// SIMATIC STEP 7 (V5.x) project EXO6
// CPU: CPU 314
// station: Matériel
// station: SIMATIC 300(1)
// station: P_ADR_BUS
// program: Programme S7(1)

SYMBOL_TABLE
"BP"	I 0.0	BOOL
"MOTEUR"	Q 0.0	BOOL
"LAMPE"	Q 0.1	BOOL
END_SYMBOL_TABLE

ORGANIZATION_BLOCK OB 1
TITLE = "Main Program Sweep (Cycle)"
VERSION : 0.1
VAR_TEMP
  OB1_EV_CLASS : BYTE ;	//Bits 0-3 = 1 (Coming event), Bits 4-7 = 1 (Event class 1)
  OB1_SCAN_1 : BYTE ;	//1 (Cold restart scan 1 of OB 1), 3 (Scan 2-n of OB 1)
  OB1_PRIORITY : BYTE ;	//Priority of OB Execution
  OB1_OB_NUMBR : BYTE ;	//1 (Organization block 1, OB1)
  OB1_RESERVED_1 : BYTE ;	//Reserved for system
  OB1_RESERVED_2 : BYTE ;	//Reserved for system
  OB1_PREV_CYCLE : INT ;	//Cycle time of previous OB1 scan (milliseconds)
  OB1_MIN_CYCLE : INT ;	//Minimum cycle time of OB1 (milliseconds)
  OB1_MAX_CYCLE : INT ;	//Maximum cycle time of OB1 (milliseconds)
  OB1_DATE_TIME : DATE_AND_TIME ;	//Date and time OB1 started
END_VAR
BEGIN
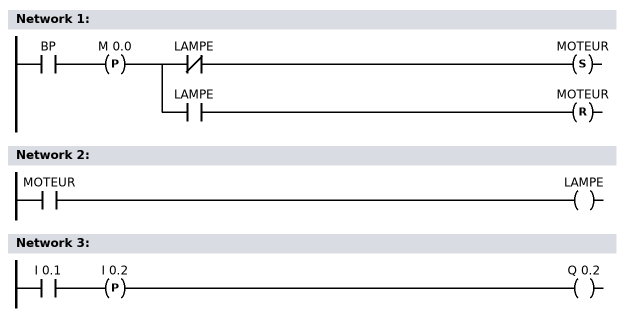
NETWORK
TITLE =
      A     "BP";
      BLD   100;
      FP    M 0.0;
      =     L 20.0;
      A     L 20.0;
      AN    "LAMPE";
      S     "MOTEUR";
      A     L 20.0;
      A     "LAMPE";
      R     "MOTEUR";
NETWORK
TITLE =
      A     "MOTEUR";
      =     "LAMPE";
NETWORK
TITLE =
      A     I 0.1;
      FP    I 0.2;
      =     Q 0.2;
NETWORK
TITLE =
END_ORGANIZATION_BLOCK
